(* IEC 61131-3 sources: JingjiangArm/moonboxpro_arm_8.4/Application/Application/任务列表/ExtTask/动作处理, 7 files *)

(* ---- CUSTOMERNAME_ENUM.st ---- *)
(*@CES
Name=CUSTOMERNAME_ENUM
Type=Gvl
TypeGuid=2db5746d-d284-4425-9f7f-2663a34b0ebc
Guid=89f6971c-faf5-49c1-98cd-d55cef9a6f12
HasDeclaration=True
HasImplementation=False
*)
{DECLARATION}
TYPE CUSTOMERNAME_ENUM :
(
	CUSTOMERNAME_KESAI				:= 0,
	CUSTOMERNAME_KESAI1				:= 2000,
	CUSTOMERNAME_BEIREN				:= 2001,
	CUSTOMERNAME_ALLOTEC			:= 2002,
	CUSTOMERNAME_DADONG				:= 2003,
	CUSTOMERNAME_SANLI				:= 2004,
	CUSTOMERNAME_HAPPYFIELD			:= 2005,
	CUSTOMERNAME_QIANGDA			:= 2006,
	CUSTOMERNAME_ALTMA				:= 2007,
	CUSTOMERNAME_CHENGBAO			:= 2008,
	CUSTOMERNAME_FANGBANG			:= 2009,
	CUSTOMERNAME_ZHONGBANG			:= 2010,
	CUSTOMERNAME_HUAFENG			:= 2011,
	CUSTOMERNAME_GUOWEI				:= 2012,(*2019.09.10.085124|Niu，j|国伟2012*)
	CUSTOMERNAME_JINGCAI			:= 2013,
	CUSTOMERNAME_BOCHUANG			:= 2014,(*2019.09.10.085124|Niu，j|博创2014*)
	CUSTOMERNAME_SHOUXIN			:= 2015,
	CUSTOMERNAME_MEIGE				:= 2016,
	CUSTOMERNAME_RUNXIN				:= 2017,
	CUSTOMERNAME_MINGCHENG			:= 2018,
	CUSTOMERNAME_JIATE				:= 2019,
	CUSTOMERNAME_QIAOXIN			:= 2020,
	CUSTOMERNAME_NBXINDA			:= 2021,
	CUSTOMERNAME_HAININGBANGDE		:= 2022,
	CUSTOMERNAME_FOSHANHONGYI		:= 2023,
	CUSTOMERNAME_DONGGUANHONGHE		:= 2024,
	CUSTOMERNAME_JIANGYINLIDA		:= 2025,(*2020.2.14.130743|江阴力达*)
	CUSTOMERNAME_LIJIACHUANG		:= 2026,(*2020.4.21.152846|汕头利佳创|*)
	CUSTOMERNAME_RUIANXINXIN		:= 2027,
(*2023.3.29.111636||新增整理全部厂家-兼容基础款所有厂家-人机已修改*)
	CUSTOMERNAME_HAININGRENMIN		:= 2028,(*海宁人民*)
	CUSTOMERNAME_WENZHKAIXU			:= 2029,(*温州凯旭*)
	CUSTOMERNAME_FOSHANHUIPUDA		:= 2030,(*佛山汇普达*)
	CUSTOMERNAME_WENZHHONGYANG		:= 2031,(*温州宏阳*)
	CUSTOMERNAME_JIANGYINHUITELI	:= 2032,(*江阴汇特力*)
	CUSTOMERNAME_WUXIHONGRUI		:= 2033,(*无锡宏瑞*)
	CUSTOMERNAME_FOSHANSHENGTU		:= 2034,(*佛山盛图*)
	CUSTOMERNAME_WEINANRENMIN		:= 2035,(*渭南人民*)
	CUSTOMERNAME_MINGDING			:= 2036,(*2022.10.19.104419|汕头铭鼎|*)
	CUSTOMERNAME_SHANTOUSHIBIAO		:= 2037,(*汕头世标*)
	CUSTOMERNAME_LINANSHENGHONG		:= 2038,(*临安盛宏*)
	CUSTOMERNAME_WEINANYIJIANGCHENG	:= 2039,(*渭南一匠成*)
	CUSTOMERNAME_ZHEJIANGDEGUANG	:= 2040,(*浙江德光*)
	CUSTOMERNAME_WEINANSHENGTAI		:= 2041,(*渭南盛泰*)
	CUSTOMERNAME_JIANGYINHUITONG	:= 2042,(*江阴汇通2022.7.7.103023*)

	CUSTOMERNAME_GAOMINGZHENGYI		:= 2043,(*高明正一*)
	CUSTOMERNAME_ZHEJIANGJINGBANG	:= 2044,(*浙江劲邦*)
	CUSTOMERNAME_DONGGUANJINKUN		:= 2045,(*东莞晋坤*)
	CUSTOMERNAME_RUIANYAOFENG		:= 2046,(*瑞安耀峰*)
	CUSTOMERNAME_WEINANJIARUI		:= 2047,(*渭南嘉瑞*)
	CUSTOMERNAME_FOSHANCHONGYUAN	:= 2048,(*佛山崇源*)
	CUSTOMERNAME_CHANGLEHUAZHOU		:= 2049,(*长乐华周*)
	CUSTOMERNAME_WEINANWODE			:= 2050,(*渭南沃德*)
	CUSTOMERNAME_XIANQINHUA			:= 2051,(*西安秦华*)
	CUSTOMERNAME_ZHEJIANGOUNUO		:= 2052,(*浙江欧诺*)
	CUSTOMERNAME_WENZHOUZHEKE		:= 2053,(*温州浙科*)
	CUSTOMERNAME_SHUNDEDELI			:= 2054,(*顺德得力*)
	CUSTOMERNAME_CHAOZHOURUILONG	:= 2055,(*潮州瑞龙*)
	(*2023.10.05.150644 增加*)
	CUSTOMERNAME_WENZHOURUIGUANG	:= 2056,(*温州瑞光印刷机械*)
	CUSTOMERNAME_RUIANHONGXIANG		:= 2057,(*瑞安市鸿翔印刷机械*)
	CUSTOMERNAME_WENZHOUZHONGYIN	:= 2058,(*温州中印印刷机械*)
	CUSTOMERNAME_YOUTAIKE			:= 2059,(*渭南优泰克印刷机械有限公司@2025.3.27.093550+*)
	CUSTOMERNAME_RUIANCHENXU		:= 2060,(*瑞安市晨旭印刷机械*)
	CUSTOMERNAME_XINHONGWU			:= 2061,(*新宏吴@2025.3.27.093600*)
	CUSTOMERNAME_YUNCHENGZHIBAN		:= 2064,(*运城制版印刷机械制造有限公司*)
	CUSTOMERNAME_QINHUA				:= 2065,(*运城制版印刷机械制造有限公司*)
	(*2023.10.05.150644 新增*)
	CUSTOMERNAME_CHAOXU				:= 2066,(*温州超旭*)

	CUSTOMERNAME_BEIREN_NOLOGO		:= 2999(*2022.7.18.154922*)
);
END_TYPE

{IMPLEMENTATION}

(* ---- GLOBALSTS_ENUMS.st ---- *)
(*@CES
Name=GLOBALSTS_ENUMS
Type=Gvl
TypeGuid=2db5746d-d284-4425-9f7f-2663a34b0ebc
Guid=72e745eb-8b64-4285-a625-315fc9f93d85
HasDeclaration=True
HasImplementation=False
*)
{DECLARATION}
TYPE GLOBALSTS_ENUMS :
(
	GSE_ESTOP				:= 1,(*急停状态|*)
	GSE_STOP				:= 2,(*停机状态|*)
	GSE_ACCING				:= 3,(*加速状态|*)
	GSE_DECING				:= 4,(*减速状态|*)
	GSE_INK					:= 5,(*空转状态|*)
	GSE_PRINT				:= 6,(*印刷状态|*)
	GSE_PRESTART			:= 7,(*预启动|*)
	GSE_KEEP_TENSION		:= 8,(*保持张力|*)
	GSE_PRINT_PRESTART		:= 9,(*印刷预启动|*)
	GSE_UNKNOWN				:= -1(*未知状态|*)
);
END_TYPE

{IMPLEMENTATION}

(* ---- StFlag_UserActCtl.st ---- *)
(*@CES
Name=StFlag_UserActCtl
Type=Gvl
TypeGuid=2db5746d-d284-4425-9f7f-2663a34b0ebc
Guid=e0d5b7fa-b2d2-412b-a1dd-76db7c909aa8
HasDeclaration=True
HasImplementation=False
*)
{DECLARATION}
TYPE StFlag_UserActCtl :
(*为了全局参数不到流程里面，将流程里用到的变量整理一个结构体把，这样简单一点*)
STRUCT
END_STRUCT
END_TYPE

{IMPLEMENTATION}

(* ---- TypEnumDataType.st ---- *)
(*@CES
Name=TypEnumDataType
Type=Gvl
TypeGuid=2db5746d-d284-4425-9f7f-2663a34b0ebc
Guid=1087113d-025e-4430-94e5-1f2f37c86e74
HasDeclaration=True
HasImplementation=False
*)
{DECLARATION}
TYPE TypEnumDataType :
(
		TYPE_LREAL,
		TYPE_REAL,
		TYPE_DINT,
		TYPE_DWORD,
		TYPE_INT,
		TYPE_WORD,
		TYPE_BYTE,
		TYPE_BOOL
);
END_TYPE

{IMPLEMENTATION}

(* ---- KS_SetVarValue_NQ0.st ---- *)
(*@CES
Name=KS_SetVarValue_NQ0
Type=FunctionBlock
TypeGuid=6f9dac99-8de1-4efc-8465-68ac443b7d08
Guid=b4c3880f-3565-4c03-a3ee-9be25f97e488
HasDeclaration=True
HasImplementation=True
*)
{DECLARATION}
FUNCTION KS_SetVarValue_NQ0 : BOOL
VAR_INPUT
	i_dwVarAdr:DWORD;(*变量地址*)
	i_iSetValue:INT;(*设置的初始值|暂定设置的初始值为int型*)
	i_EmVarType:TypEnumDataType;(*变量类型*)
END_VAR
VAR
	piVar:POINTER TO INT;
END_VAR
{IMPLEMENTATION}
IF i_dwVarAdr<>0 THEN;ELSE RETURN;END_IF
CASE i_EmVarType OF
TYPE_BOOL:;
TYPE_INT:
	piVar:=i_dwVarAdr;
	IF piVar^=0 THEN
		piVar^:=i_iSetValue;
	END_IF
TYPE_WORD:;
TYPE_DWORD:;
TYPE_REAL:;
TYPE_LREAL:;
ELSE;
END_CASE

(* ---- KS_FB_BlowerFunction.st ---- *)
(*@CES
Name=KS_FB_BlowerFunction
Type=FunctionBlock
TypeGuid=6f9dac99-8de1-4efc-8465-68ac443b7d08
Guid=d1a93ad3-e4c3-4af6-9dda-58720c2c75d3
HasDeclaration=True
HasImplementation=True
*)
{DECLARATION}
FUNCTION_BLOCK KS_FB_BlowerFunction
VAR_INPUT
	i_xEn					:BOOL;(*功能使能*)
	i_xAllStartOrStop_Trig	:BOOL;(*全体启动或者停止|沿触发|延时启动*)
	i_xStartByKnob			:BOOL;(*单轴启动根据旋钮开关标志|用于开关控制启动的逻辑|无则不输入*)
	i_iAllStartDelayTime	:INT;(*全体启动延时S*)
	i_iCycleTime_Plc		:INT;(*程序执行时间*)
	i_iAxisSum				:INT;(*轴总数*)
	i_paiAxisNumList		:POINTER TO ARRAY [1..MAX_UNIT_NUM] OF INT;(*轴号列表*)
	i_paxAxisStartEn		:POINTER TO ARRAY [1..MAX_UNIT_NUM] OF BOOL;(*轴启动使能|有效后按钮开关才能起作用*)
	i_paxStartKnob			:POINTER TO ARRAY [1..MAX_UNIT_NUM] OF BOOL;(*全体启动,每个轴旋钮输入*)
	i_paxStartOrStopBtn		:POINTER TO ARRAY [1..MAX_UNIT_NUM] OF BOOL;(*单轴的启动停止按钮*)
	i_paxNeedStop			:POINTER TO ARRAY [1..MAX_UNIT_NUM] OF BOOL;(*单轴需要停止输出标志*)
	i_paxAxisStarted		:POINTER TO ARRAY [1..MAX_UNIT_NUM] OF BOOL;(*单个轴的启动输出标志|实际处于启动状态，
																			可以根据i_paxNeedStop这个变量控制实际输出*)
END_VAR
VAR_OUTPUT
	o_xEn:BOOL;
	o_xAllStarted:BOOL;(*全体启动标志*)
	o_xAutoStartDne:BOOL;(*自动启动轴启动完成*)
	o_iStartedSum:INT;(*启动的总数*)
END_VAR
VAR
	iN: INT;
	xEned: BOOL;(*进入过使能状态*)
	iAxisNum: INT;(*轴号*)
	xPreAllStartOrStop_Trig: BOOL;(*全部启动或者停止上个周期标志*)
	axAllStartedTemp:ARRAY [1..MAX_UNIT_NUM] OF BOOL;(*单个轴的启动了*)
	axAutoStarted: ARRAY [1..MAX_UNIT_NUM] OF BOOL;(*自动启动的标志*)
	axPreStartOrStopBtn: ARRAY [1..MAX_UNIT_NUM] OF BOOL;(*手动按钮由于沿处理标志*)
	xTimeUp: BOOL;(*计时时间到*)
	iCnt: INT;(*计数值*)
	(*旋钮取沿|用于旋钮控制启动停止方式*)
	afbKnobRTrig: ARRAY [1..MAX_UNIT_NUM] OF R_TRIG;
	afbKnobFTrig: ARRAY [1..MAX_UNIT_NUM] OF F_TRIG;
END_VAR

{IMPLEMENTATION}
IF i_paxStartKnob<>0 AND
	i_paxNeedStop<>0 AND
 	i_paxStartOrStopBtn<>0 AND
	i_paxAxisStartEn<>0 AND
	i_paiAxisNumList<>0 AND
	i_paxAxisStarted<>0 THEN

	IF i_iCycleTime_Plc<=0 THEN
		i_iCycleTime_Plc:=gc_EXT_TSK_CYCLE_TIME;
	END_IF

	IF i_xEn THEN
		(*旋钮控制*)
		IF i_xStartByKnob THEN(*根据旋钮状态控制|按钮将不起作用*)
			o_xAllStarted:=FALSE;
			FOR iN:=1 TO i_iAxisSum BY 1 DO
				iAxisNum:=i_paiAxisNumList^[iN];
				IF iAxisNum>0 AND iAxisNum<=MAX_UNIT_NUM THEN;
					afbKnobRTrig[iAxisNum](CLK:=i_paxStartKnob^[iAxisNum]);
					afbKnobFTrig[iAxisNum](CLK:=i_paxStartKnob^[iAxisNum]);
					IF afbKnobRTrig[iAxisNum].Q THEN
						axAllStartedTemp[iAxisNum]:=TRUE;
					ELSIF afbKnobFTrig[iAxisNum].Q THEN
						axAllStartedTemp[iAxisNum]:=FALSE;
					END_IF
				END_IF
			END_FOR
		ELSE
(*--------------------------自动部分START-------------------------*)
			xTimeUp:=FALSE;
			(*全体启动部分*)
			IF  i_xAllStartOrStop_Trig AND NOT xPreAllStartOrStop_Trig THEN(*启动按键按下*)
				o_xAllStarted:=NOT o_xAllStarted;
				IF o_xAllStarted THEN(*启动了|清零周期计数|并输出时间到标志打开第一个轴*)
					iCnt:=0;
					xTimeUp:=TRUE;
				END_IF
			END_IF

			(*计时部分*)
			iCnt:=iCnt+1;
			IF o_xAutoStartDne THEN(*自动启动完成后清零计数值*)
				iCnt:=0;
			END_IF
			IF iCnt>i_iAllStartDelayTime*1000/i_iCycleTime_Plc THEN(*时间到*)
				iCnt:=0;
				xTimeUp:=TRUE;
			END_IF

			(*自动控制延时启动*)
			FOR iN:=1 TO i_iAxisSum BY 1 DO
				iAxisNum:=i_paiAxisNumList^[iN];
				IF iAxisNum>0 AND iAxisNum<=MAX_UNIT_NUM THEN(*轴号是否合法*)
					IF o_xAllStarted THEN(*全体启动了|延时启动|只自动启动一次*)
						IF i_paxStartKnob^[iAxisNum] AND i_paxAxisStartEn^[iAxisNum] THEN(*开关打开了*)
							IF NOT axAutoStarted[iAxisNum]  THEN(*未自动启动*)
								IF NOT axAllStartedTemp[iAxisNum] THEN(*未启动*)
									IF xTimeUp THEN(*计时到了*)
										axAllStartedTemp[iAxisNum]:=TRUE;
										axAutoStarted[iAxisNum]:=TRUE;
										xTimeUp:=FALSE;
									END_IF
								ELSE
									axAutoStarted[iAxisNum]:=TRUE;
								END_IF
							END_IF
						END_IF
					END_IF

					IF (NOT o_xAllStarted OR
						NOT i_paxStartKnob^[iAxisNum] OR
						NOT i_paxAxisStartEn^[iAxisNum])AND
						axAutoStarted[iAxisNum] THEN(*已经自动打开了|我们关闭它*)
						axAllStartedTemp[iAxisNum]:=FALSE;
						axAutoStarted[iAxisNum]:=FALSE;
					END_IF
				END_IF
			END_FOR

			(*查看自动启动是否完成*)
			o_xAutoStartDne:=TRUE;
			IF o_xAllStarted THEN(*全体启动了*)
				FOR iN:=1 TO i_iAxisSum BY 1 DO
					iAxisNum:=i_paiAxisNumList^[iN];
					IF i_paxStartKnob^[iAxisNum] AND
						i_paxAxisStartEn^[iAxisNum] AND
						NOT axAutoStarted[iAxisNum] THEN
						o_xAutoStartDne:=FALSE;
						EXIT;
					ELSE;
					END_IF
				END_FOR
			END_IF
(*--------------------------自动部分END-------------------------*)
		END_IF

(*--------------------------手动部分START-------------------------*)
		(*手动控制按钮启动停止部分*)
		FOR iN:=1 TO i_iAxisSum BY 1 DO
			iAxisNum:=i_paiAxisNumList^[iN];
			IF i_paxStartOrStopBtn^[iAxisNum] AND
				NOT axPreStartOrStopBtn[iAxisNum] THEN(*按下按钮*)
				axAllStartedTemp[iAxisNum]:=NOT axAllStartedTemp[iAxisNum];
			END_IF

			(*在这个循环里面处理轴启动使能标志对输出的影响*)
			IF NOT i_paxAxisStartEn^[iAxisNum] THEN;
				axAllStartedTemp[iAxisNum]:=FALSE;
			END_IF
		END_FOR
(*--------------------------手动部分END-------------------------*)
		xEned:=TRUE;
	ELSE(*功能块未使能*)
		IF xEned THEN
			xEned:=FALSE;
			o_xAllStarted:=FALSE;
			o_xAutoStartDne:=FALSE;
			FOR  iN:=1 TO i_iAxisSum BY 1 DO
				iAxisNum:=i_paiAxisNumList^[iN];
				IF iAxisNum>0 AND iAxisNum<=MAX_UNIT_NUM THEN
					axAllStartedTemp[iAxisNum]:=FALSE;
					axAutoStarted[iAxisNum]:= FALSE(*TRUE*); (* 2021.3.31.092022/参照2021.3.32在欧泰715机器上更新(汕头彭城) *)
				END_IF
			END_FOR
		END_IF
	END_IF

	(*最终输出控制*)
	o_iStartedSum:=0;
	FOR  iN:=1 TO i_iAxisSum BY 1 DO
		iAxisNum:=i_paiAxisNumList^[iN];
		i_paxAxisStarted^[iAxisNum]:=axAllStartedTemp[iAxisNum];
		IF i_paxNeedStop^[iAxisNum] THEN
			i_paxAxisStarted^[iAxisNum]:=FALSE;
		END_IF

		(*统计实际输出的个数*)
		IF i_paxAxisStarted^[iAxisNum] THEN
			o_iStartedSum:=o_iStartedSum+1;
		END_IF

		(* 2020.11.3.110550|lyt|修复已知的bug *)
		axPreStartOrStopBtn[iAxisNum]:=i_paxStartOrStopBtn^[iAxisNum];
	END_FOR

	xPreAllStartOrStop_Trig:=i_xAllStartOrStop_Trig;
END_IF
o_xEn:=i_xEn;

(* ---- KS_FB_GrpLampAndAlarmBellCtl.st ---- *)
(*@CES
Name=KS_FB_GrpLampAndAlarmBellCtl
Type=FunctionBlock
TypeGuid=6f9dac99-8de1-4efc-8465-68ac443b7d08
Guid=eea8cc40-7b3e-4264-b59d-3f431f7baf96
HasDeclaration=True
HasImplementation=True
*)
{DECLARATION}
FUNCTION_BLOCK KS_FB_GrpLampAndAlarmBellCtl
VAR_INPUT
	i_xEn: BOOL;
	i_iUnitNum: INT;
	i_pstStEvtReq: POINTER TO StEvtReq;
	i_xFlag_Stoping: BOOL;
	i_xFlag_Stop: BOOL;
END_VAR
VAR_OUTPUT
	o_xEn: BOOL;
	o_iErNo: INT;
END_VAR
VAR
	tmNow: TIME;
	tmLastStateChanged_Stop: TIME;
	xLamp_Stop: BOOL;(*停止指示灯*)
END_VAR

{IMPLEMENTATION}
o_xEn:= i_xEn;
o_iErNo:= 0;
IF i_xEn THEN
	tmNow:= TIME();
	IF i_xFlag_Stoping THEN(*停机过程中停止指示灯闪烁*)
		IF tmNow-tmLastStateChanged_Stop>=T#200MS THEN
			xLamp_Stop:= NOT xLamp_Stop;
			tmLastStateChanged_Stop:= tmNow;
		END_IF
	ELSE
		xLamp_Stop:= i_xFlag_Stop;
		tmLastStateChanged_Stop:= tmNow;
	END_IF

ELSE
	o_iErNo:= -1;
END_IF
